(* IEC 61131-3 sources: plc-vscode/tests/st/test-ready/trust-platform/crates/trust-runtime/tests/fixtures/plcopen_motion/single_axis_negative_public_surface/src, 2 files *)

(* ---- main.st ---- *)
PROGRAM Main
VAR
    WrongError : MC_ERROR;
    WrongPayload : MC_PAYLOAD_REF;
END_VAR
END_PROGRAM

(* ---- tests.st ---- *)
TEST_PROGRAM plcopen_motion_single_axis_negative_public_surface
VAR
    WrongError : MC_ERROR;
    WrongPayload : MC_PAYLOAD_REF;
END_VAR
END_TEST_PROGRAM
